Fanuc KAREL source: kt00888.KL

-- PROVISIONAL review KL for V1013-1; original PC SHA256 c53f3fa47288e39b1d27833a5729c8b59453af1f9f0d23a259f21d81d127c4b6
-- Incomplete behavior may be omitted. Consult companion uncertainty JSON. Do not deploy.
PROGRAM KT00888
%NOLOCKGROUP
-- UNRESOLVED_DECL P1 type=000101
-- UNRESOLVED_DECL P2 type=000101
-- UNRESOLVED_DECL OUT type=000101
BEGIN
  -- UNRESOLVED_PC offsets 5-32; opcodes 27,22,1C,76,7E,4A
  -- UNRESOLVED_PC offsets 37-41; opcodes 7F
END KT00888
